Fanuc KAREL source: kt00024.KL

-- PROVISIONAL review KL for V1013-1; original PC SHA256 b07fb6cb7d50188418c340196d7c61d4cffe0e04b3c8ba1b59bec42e6b798298
-- Incomplete behavior may be omitted. Consult companion uncertainty JSON. Do not deploy.
PROGRAM KT00024
%NOLOCKGROUP
VAR
  OUT : REAL
-- UNRESOLVED_DECL Y1 type=002018
-- UNRESOLVED_DECL H2 type=002017
BEGIN
  -- UNRESOLVED_PC offsets 5-19; opcodes 2E,22,9D,33,B2
  -- UNRESOLVED_PC offsets 24-38; opcodes 2E,22,9D,33,B4
  -- UNRESOLVED_PC offsets 43-69; opcodes 22,9D,33,B1,22,9D,33,B3,52,64,23
  -- UNRESOLVED_PC offsets 74-78; opcodes 7F
END KT00024
